// TIA Portal project "GARAJ OTOMASYONU" (V18)

(* hardware
DEVICE "S7-1200 station_1"  S7-1200 Station
   slot 0: "Rack_0"  S7-1200 Rack  Rack  V1.0
   slot 1: "PLC_1"  CPU 1214C AC/DC/Rly  6ES7 214-1BG40-0XB0  V4.6
*)

// ===== PLC "PLC_1"  CPU 1214C AC/DC/Rly =====

VAR_GLOBAL   // PLC tag table "Default tag table"
   "MAN-OTO ANAHTARI" AT %I0.0 : Bool;
   "MAN AC BUT" AT %I0.1 : Bool;
   "MAN KAPAT BUT" AT %I0.2 : Bool;
   "FOTOSEL 1" AT %I0.3 : Bool;
   "FOTOSEL 2" AT %I0.4 : Bool;
   "KAPI ACIK SWITCH" AT %I0.5 : Bool;
   "KAPI KAPALI SWITCH" AT %I0.6 : Bool;
   "KAPI ACMA VALFI" AT %Q0.0 : Bool;
   "KAPI KAPATMA VALFI" AT %Q0.1 : Bool;
   "OTO CALISMA MEM" AT %M10.0 : Bool;
   "MAN AC MEM" AT %M10.1 : Bool;
   "MAN KAPAT MEM" AT %M10.2 : Bool;
   "OTO AC MEM" AT %M10.3 : Bool;
   "OTO KAPAT MEM" AT %M10.4 : Bool;
END_VAR

// folder: System blocks/Program resources

DATA_BLOCK "TIMER 1"   // DB1
{ S7_Optimized_Access := 'TRUE' }
AUTHOR : Simatic
FAMILY : IEC
NAME : IEC_TMR
VERSION : 1.0
// stored: InstanceOfName IEC_TIMER
"IEC_TIMER"
BEGIN
END_DATA_BLOCK

// folder: (top level)

ORGANIZATION_BLOCK "Main"   // OB1, LAD, ProgramCycle
TITLE = "Main Program Sweep (Cycle)"
{ S7_Optimized_Access := 'TRUE' }
VERSION : 0.1
   VAR_INPUT
      Initial_Call : Bool;   // Initial call of this OB
      Remanence : Bool;   // =True, if remanent data are available
   END_VAR
BEGIN

REGION Network 1: MANUEL-OTOMATIK CALISMA SECIMI
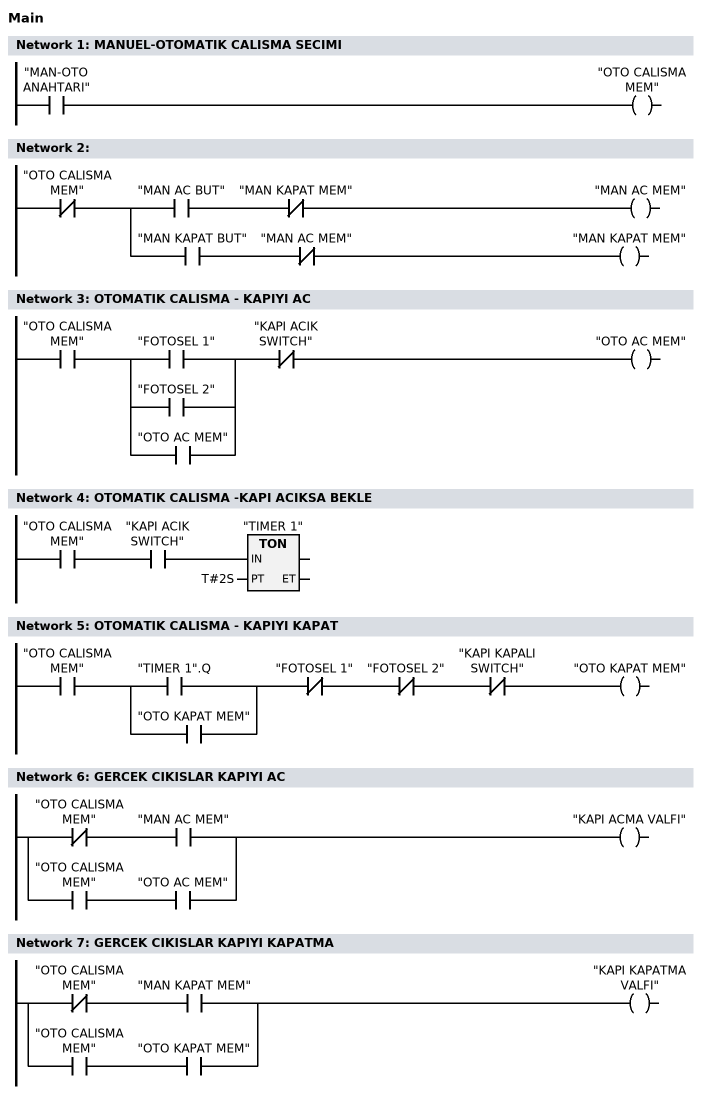
   RUNG wire#powerrail
      Contact( "MAN-OTO ANAHTARI" )
      Coil( "OTO CALISMA MEM" )
   END_RUNG
   // the same network as SCL:
   "OTO CALISMA MEM" := "MAN-OTO ANAHTARI";
END_REGION

REGION Network 2
   RUNG wire#powerrail
      I_Contact( "OTO CALISMA MEM" )
      wire#w1
      Contact( "MAN AC BUT" )
      I_Contact( "MAN KAPAT MEM" )
      Coil( "MAN AC MEM" )
   END_RUNG
   RUNG wire#w1
      Contact( "MAN KAPAT BUT" )
      I_Contact( "MAN AC MEM" )
      Coil( "MAN KAPAT MEM" )
   END_RUNG
   // the same network as SCL:
   "MAN AC MEM" := NOT "OTO CALISMA MEM" AND "MAN AC BUT" AND NOT "MAN KAPAT MEM";
   "MAN KAPAT MEM" := NOT "OTO CALISMA MEM" AND "MAN KAPAT BUT" AND NOT "MAN AC MEM";
END_REGION

REGION Network 3: OTOMATIK CALISMA - KAPIYI AC
   RUNG wire#powerrail
      Contact( "OTO CALISMA MEM" )
      wire#w1
      Contact( "FOTOSEL 1" )
      wire#w2
      I_Contact( "KAPI ACIK SWITCH" )
      Coil( "OTO AC MEM" )
   END_RUNG
   RUNG wire#w1
      Contact( "FOTOSEL 2" )
   END_RUNG wire#w2
   RUNG wire#w1
      Contact( "OTO AC MEM" )
   END_RUNG wire#w2
   // the same network as SCL:
   "OTO AC MEM" := "OTO CALISMA MEM" AND ("FOTOSEL 1" OR "FOTOSEL 2" OR "OTO AC MEM") AND NOT "KAPI ACIK SWITCH";
END_REGION

REGION Network 4: OTOMATIK CALISMA -KAPI ACIKSA BEKLE
   "TIMER 1".TON(IN := "OTO CALISMA MEM" AND "KAPI ACIK SWITCH", PT := T#2S);
END_REGION

REGION Network 5: OTOMATIK CALISMA - KAPIYI KAPAT
   RUNG wire#powerrail
      Contact( "OTO CALISMA MEM" )
      wire#w1
      Contact( "TIMER 1".Q )
      wire#w2
      I_Contact( "FOTOSEL 1" )
      I_Contact( "FOTOSEL 2" )
      I_Contact( "KAPI KAPALI SWITCH" )
      Coil( "OTO KAPAT MEM" )
   END_RUNG
   RUNG wire#w1
      Contact( "OTO KAPAT MEM" )
   END_RUNG wire#w2
   // the same network as SCL:
   "OTO KAPAT MEM" := "OTO CALISMA MEM" AND ("TIMER 1".Q OR "OTO KAPAT MEM") AND NOT "FOTOSEL 1" AND NOT "FOTOSEL 2" AND NOT "KAPI KAPALI SWITCH";
END_REGION

REGION Network 6: GERCEK CIKISLAR KAPIYI AC
   RUNG wire#powerrail
      I_Contact( "OTO CALISMA MEM" )
      Contact( "MAN AC MEM" )
      wire#w1
      Coil( "KAPI ACMA VALFI" )
   END_RUNG
   RUNG wire#powerrail
      Contact( "OTO CALISMA MEM" )
      Contact( "OTO AC MEM" )
   END_RUNG wire#w1
   // the same network as SCL:
   "KAPI ACMA VALFI" := (NOT "OTO CALISMA MEM" AND "MAN AC MEM") OR ("OTO CALISMA MEM" AND "OTO AC MEM");
END_REGION

REGION Network 7: GERCEK CIKISLAR KAPIYI KAPATMA
   RUNG wire#powerrail
      I_Contact( "OTO CALISMA MEM" )
      Contact( "MAN KAPAT MEM" )
      wire#w1
      Coil( "KAPI KAPATMA VALFI" )
   END_RUNG
   RUNG wire#powerrail
      Contact( "OTO CALISMA MEM" )
      Contact( "OTO KAPAT MEM" )
   END_RUNG wire#w1
   // the same network as SCL:
   "KAPI KAPATMA VALFI" := (NOT "OTO CALISMA MEM" AND "MAN KAPAT MEM") OR ("OTO CALISMA MEM" AND "OTO KAPAT MEM");
END_REGION
END_ORGANIZATION_BLOCK